Fanuc KAREL source: KT00847.KL

PROGRAM KT00847
%NOLOCKGROUP
VAR
  R1: REAL
  R2: REAL
  OUT: REAL
BEGIN
  R1 = 2.0
  R2 = 3.0
  R1 = 2.0
  R2 = 3.0
  OUT = TAN(R1)
END KT00847
